TYPE ST_PhysicalOutputs :
STRUCT
    bSafetyRunRequest                  : BOOL;
    bSafetyResetRequest                : BOOL;
    bSafetyErrorAcknowledgementRequest : BOOL;
    bAirSupplyEnable                   : BOOL;
    bMainDoorLockRequest               : BOOL;
    bIndexRotatePortA                  : BOOL;
    bIndexStopPortB                    : BOOL;
    bLedStart                          : BOOL;
    bLedReset                          : BOOL;
    bStatusIndicator                  : BOOL;
    bInternalLight                    : BOOL;
    bNestLight                        : BOOL;
END_STRUCT
END_TYPE

(* stored: Version 1.1.0.1, ProductVersion 3.1.4026.18
   DUT ST_PhysicalOutputs: Id {c6982397-4202-4d85-945a-2aa8bb403ca0} *)
